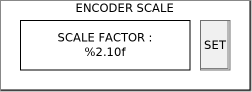
VISUALIZATION ENCODER  // 252x92
    Rectangle (0,0 250x90), "ENCODER SCALE"
    Rectangle (20,20 170x50), "SCALE FACTOR : %2.10f", text variable: MAIN.Track.EncoderScalingFactor
        OnMouseDown: write the text variable via VisuDialogs.Numpad, title 'Scaling Factor'
    Button (200,20 30x50), "SET"
        tap MAIN.Track.EncoderReset
END_VISUALIZATION

(* stored: Version 1.1.0.1, ProductVersion 3.1.4024.16
   Visu ENCODER: Id {34e6ee01-cca1-4aa5-8dd7-b1e006bb2f9f} *)
